Fanuc KAREL source: KD00049.KL

PROGRAM KD00049
%NOLOCKGROUP
%DEFGROUP = 1
VAR
  I: INTEGER
  J: INTEGER
  B: BOOLEAN
  R: REAL
  S: STRING[80]
BEGIN
  MOVE AWAY 10.0
END KD00049
